RoboDK station: RobodkBasico-2.rdk

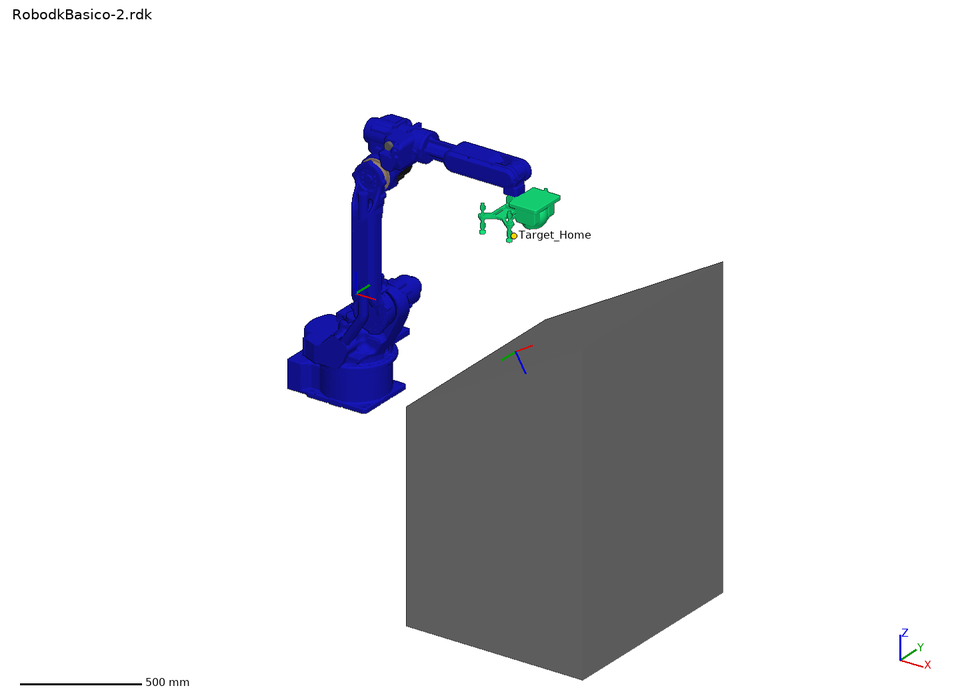
[picture v0: the station drawn from its stored meshes, robots at their saved joint values, targets as dots, program paths as lines]
Station RobodkBasico-2 (saved by RoboDK 6.0.6). Poses are relative to the parent item; angles as X-Y-Z fixed-axis rotations.
Station parameters (name, value as stored): LIN64
  - frame Motoman MH6 Base at (0, 0, 450) mm
    - robot Motoman MH6: 6 axes, payload 6 kg, reach 1422 mm, repeatability 0.08 mm, weight 130 kg
        modified DH rows (alpha deg, a mm, theta deg, d mm): 0, 0, 0, 450; -90, 152, -90, 0; 0, 614, 0, 0; -90, 155, 0, 640; 90, 0, 90, 0; -90, 0, 0, 95
        base shift (0, 0, -450) mm
        joint limits [-170, -90, -175, -180, -45, -360] to [170, 155, 250, 180, 225, 360]; home [0, 0, 0, 0, 0, 0]; saved at [0, 0, 0, 0, 0, 0]
      - tool Ventosas, TCP at (0, 0, 190) mm, size 250 x 290 x 148 mm
    - frame Frame_from_Target1 at (823.2, -34.49, -21.13) mm, rotated rx -180 ry -30 rz 0 deg
      - target Target_Home (Cartesian target) at (225.55, -34.49, -453.06) mm, rotated rx 0 ry -30 rz 0 deg; joints [0, 0, 0, 0, 0, 0] of Motoman MH6
  - object CAJA2 at (1600, 500, 300) mm, rotated rx 180 ry 0 rz 0 deg, size 886.4 x 1000 x 1511.7 mm, geometry from CAJA2.stp
  - Python program RosPolar (listed below)
  - Python program Trébol (listed below)
  - Python program Elipse (listed below)

--- Python program RosPolar ---
from robodk.robolink import *    # API para comunicarte con RoboDK
from robodk.robomath import *    # Funciones matemáticas
import math
from matplotlib.textpath import TextPath
from matplotlib.path import Path
#------------------------------------------------
# 1) Conexión a RoboDK e inicialización
#------------------------------------------------
RDK = Robolink()

# Elegir un robot (si hay varios, aparece un popup)
robot = RDK.ItemUserPick("Selecciona un robot", ITEM_TYPE_ROBOT)
if not robot.Valid():
    raise Exception("No se ha seleccionado un robot válido.")

### Conectar al robot físico
##if not robot.Connect():
##    raise Exception("No se pudo conectar al robot. Verifica que esté en modo remoto y que la configuración sea correcta.")
##
### Confirmar conexión
##if not robot.ConnectedState():
##    raise Exception("El robot no está conectado correctamente. Revisa la conexión.")
##
##print("Robot conectado correctamente.")

#------------------------------------------------
# 2) Cargar el Frame (ya existente) donde quieres dibujar
#    Ajusta el nombre si tu Frame se llama diferente
#------------------------------------------------
frame_name = "Frame_from_Target1"
frame = RDK.Item(frame_name, ITEM_TYPE_FRAME)
if not frame.Valid():
    raise Exception(f'No se encontró el Frame "{frame_name}" en la estación.')

target_name = "Target_Home"
target = RDK.Item(target_name , ITEM_TYPE_TARGET)
if not target.Valid():
    print(f"Error: El target '{target_name}' no existe en la estación.")

# Asignamos este frame al robot
robot.setPoseFrame(frame)
# Usamos la herramienta activa
robot.setPoseTool(robot.PoseTool())

# Ajustes de velocidad y blending
robot.setSpeed(300)   # mm/s - Ajusta según necesites
robot.setRounding(5)  # blending (radio de curvatura)

#------------------------------------------------
# 3) Parámetros de la figura (rosa polar)
#------------------------------------------------
num_points = 100      # Cuántos puntos muestreamos (mayor = más suave)
a = 60
b = 6
z_surface = 0          # Z=0 en el plano del frame
z_safe = 50            # Altura segura para aproximarse y salir

path_jose = TextPath((0, 0), "Jose", size=50)
path_leonardo = TextPath((0, -50), "Leonardo", size=50)

path = Path.make_compound_path(path_jose, path_leonardo)
puntos = path.vertices
instrucciones = path.codes

#------------------------------------------------
# 4) Movimiento al centro en altura segura
#------------------------------------------------
# El centro de la rosa (r=0) corresponde a x=0, y=0
robot.MoveJ(target)
robot.MoveJ(transl(0, 0, z_surface - z_safe))

# Bajamos a la "superficie" (Z=0)
robot.MoveL(transl(0, 0, z_surface))

# #------------------------------------------------
# # 5) Dibujar la rosa polar
# #    r = a - b*cos(theta)
# #    x = r*cos(theta), y = r*sin(theta)
# #------------------------------------------------
# # Recorremos theta de 0 a 2*pi (una vuelta completa)
# full_turn = 2*math.pi

# for i in range(num_points+1):
#     # Fracción entre 0 y 1
#     t = i / num_points
#     # Ángulo actual
#     theta = full_turn * t

#     # Calculamos r
#     r = a - b*math.cos(theta)

#     # Convertimos a coordenadas Cartesianas X, Y
#     x = r * math.cos(theta)
#     y = r * math.sin(theta)

#     # Movemos linealmente (MoveL) en el plano del Frame
#     robot.MoveL(transl(x, y, z_surface))

# # Al terminar, subimos de nuevo para no chocar
# robot.MoveL(transl(x, y, z_surface - z_safe))
# robot.MoveL(target)


# #------------------------------------------------
# # 5) Dibujar la elipse
# #    r = ab/sqrt((b*cos(theta))^2 + (a*sin(theta))^2)
# #    x = r*cos(theta), y = r*sin(theta)
# #------------------------------------------------
# # Recorremos theta de 0 a 2*pi (una vuelta completa)
# full_turn = 2*math.pi

# for i in range(num_points+1):
#     # Fracción entre 0 y 1
#     t = i / num_points
#     # Ángulo actual
#     theta = full_turn * t

#     # Calculamos r
#     r = a*b/sqrt((b*math.cos(theta))**2 + (a*math.sin(theta))**2)

#     # Convertimos a coordenadas Cartesianas X, Y
#     x = r * math.cos(theta)
#     y = r * math.sin(theta)

#     # Movemos linealmente (MoveL) en el plano del Frame
#     robot.MoveL(transl(x, y, z_surface))

# # Al terminar, subimos de nuevo para no chocar
# robot.MoveL(transl(x, y, z_surface - z_safe))
# robot.MoveL(target)

#------------------------------------------------
# 5) Dibujar la trebol b lúbulos
#    r = a*cos(b*theta)
#    x = r*cos(theta), y = r*sin(theta)
#------------------------------------------------
# Recorremos theta de 0 a 2*pi (una vuelta completa)
full_turn = 2*math.pi

for i in range(num_points+1):
    # Fracción entre 0 y 1
    t = i / num_points
    # Ángulo actual
    theta = full_turn * t

    # Calculamos r
    r = a*math.cos(b*theta)-math.cos(theta**2)

    # Convertimos a coordenadas Cartesianas X, Y
    x = r * math.cos(theta)
    y = r * math.sin(theta)

    # Movemos linealmente (MoveL) en el plano del Frame
    robot.MoveL(transl(x, y, z_surface))

# Al terminar, subimos de nuevo para no chocar
robot.MoveL(transl(x, y, z_surface - z_safe))
robot.MoveL(target)


robot.MoveL(transl(150,0,0))
robot.MoveL(transl(0,0,z_surface))

for pt, code in zip(puntos, instrucciones):
    x = pt[1]
    y = pt[0]

    if code == 1:
        # Mover por arriba en el aire y bajar el lápiz
        robot.MoveL(transl(x+150, y, z_surface + z_safe))
        robot.MoveL(transl(x+150, y, z_surface))
    else:
        # Trazo continuo de la letra sobre la superficie
        robot.MoveL(transl(x+150, y, z_surface))

robot.MoveL(transl(x, y, z_surface - z_safe))
robot.MoveJ(target)
print(f"¡Figura (rosa polar) completada en el frame '{frame_name}'!")

--- Python program Trébol ---
from robodk.robolink import *    # API para comunicarte con RoboDK
from robodk.robomath import *    # Funciones matemáticas
import math
from matplotlib.textpath import TextPath
from matplotlib.path import Path
#------------------------------------------------
# 1) Conexión a RoboDK e inicialización
#------------------------------------------------
RDK = Robolink()

# Elegir un robot (si hay varios, aparece un popup)
robot = RDK.ItemUserPick("Selecciona un robot", ITEM_TYPE_ROBOT)
if not robot.Valid():
    raise Exception("No se ha seleccionado un robot válido.")

### Conectar al robot físico
##if not robot.Connect():
##    raise Exception("No se pudo conectar al robot. Verifica que esté en modo remoto y que la configuración sea correcta.")
##
### Confirmar conexión
##if not robot.ConnectedState():
##    raise Exception("El robot no está conectado correctamente. Revisa la conexión.")
##
##print("Robot conectado correctamente.")

#------------------------------------------------
# 2) Cargar el Frame (ya existente) donde quieres dibujar
#    Ajusta el nombre si tu Frame se llama diferente
#------------------------------------------------
frame_name = "Frame_from_Target1"
frame = RDK.Item(frame_name, ITEM_TYPE_FRAME)
if not frame.Valid():
    raise Exception(f'No se encontró el Frame "{frame_name}" en la estación.')

target_name = "Target_Home"
target = RDK.Item(target_name , ITEM_TYPE_TARGET)
if not target.Valid():
    print(f"Error: El target '{target_name}' no existe en la estación.")

# Asignamos este frame al robot
robot.setPoseFrame(frame)
# Usamos la herramienta activa
robot.setPoseTool(robot.PoseTool())

# Ajustes de velocidad y blending
robot.setSpeed(300)   # mm/s - Ajusta según necesites
robot.setRounding(5)  # blending (radio de curvatura)

#------------------------------------------------
# 3) Parámetros de la figura (rosa polar)
#------------------------------------------------
num_points = 100      # Cuántos puntos muestreamos (mayor = más suave)
a = 60
b = 6
z_surface = 0          # Z=0 en el plano del frame
z_safe = 50            # Altura segura para aproximarse y salir

path_jose = TextPath((0, 0), "Jose", size=50)
path_leonardo = TextPath((0, -50), "Leonardo", size=50)

path = Path.make_compound_path(path_jose, path_leonardo)
puntos = path.vertices
instrucciones = path.codes


#------------------------------------------------
# 4) Movimiento al centro en altura segura
#------------------------------------------------
# El centro de la rosa (r=0) corresponde a x=0, y=0
robot.MoveJ(target)
robot.MoveJ(transl(0, 0, z_surface - z_safe))

# Bajamos a la "superficie" (Z=0)
robot.MoveL(transl(0, 0, z_surface))

# #------------------------------------------------
# # 5) Dibujar la rosa polar
# #    r = a - b*cos(theta)
# #    x = r*cos(theta), y = r*sin(theta)
# #------------------------------------------------
# # Recorremos theta de 0 a 2*pi (una vuelta completa)
# full_turn = 2*math.pi

# for i in range(num_points+1):
#     # Fracción entre 0 y 1
#     t = i / num_points
#     # Ángulo actual
#     theta = full_turn * t

#     # Calculamos r
#     r = a - b*math.cos(theta)

#     # Convertimos a coordenadas Cartesianas X, Y
#     x = r * math.cos(theta)
#     y = r * math.sin(theta)

#     # Movemos linealmente (MoveL) en el plano del Frame
#     robot.MoveL(transl(x, y, z_surface))

# # Al terminar, subimos de nuevo para no chocar
# robot.MoveL(transl(x, y, z_surface - z_safe))
# robot.MoveL(target)


# #------------------------------------------------
# # 5) Dibujar la elipse
# #    r = ab/sqrt((b*cos(theta))^2 + (a*sin(theta))^2)
# #    x = r*cos(theta), y = r*sin(theta)
# #------------------------------------------------
# # Recorremos theta de 0 a 2*pi (una vuelta completa)
# full_turn = 2*math.pi

# for i in range(num_points+1):
#     # Fracción entre 0 y 1
#     t = i / num_points
#     # Ángulo actual
#     theta = full_turn * t

#     # Calculamos r
#     r = a*b/sqrt((b*math.cos(theta))**2 + (a*math.sin(theta))**2)

#     # Convertimos a coordenadas Cartesianas X, Y
#     x = r * math.cos(theta)
#     y = r * math.sin(theta)

#     # Movemos linealmente (MoveL) en el plano del Frame
#     robot.MoveL(transl(x, y, z_surface))

# # Al terminar, subimos de nuevo para no chocar
# robot.MoveL(transl(x, y, z_surface - z_safe))
# robot.MoveL(target)

#------------------------------------------------
# 5) Dibujar la trebol b lúbulos
#    r = a*cos(b*theta)
#    x = r*cos(theta), y = r*sin(theta)
#------------------------------------------------
# Recorremos theta de 0 a 2*pi (una vuelta completa)
full_turn = 2*math.pi

for i in range(num_points+1):
    # Fracción entre 0 y 1
    t = i / num_points
    # Ángulo actual
    theta = full_turn * t

    # Calculamos r
    r = a*math.cos(b*theta)

    # Convertimos a coordenadas Cartesianas X, Y
    x = r * math.cos(theta)
    y = r * math.sin(theta)

    # Movemos linealmente (MoveL) en el plano del Frame
    robot.MoveL(transl(x, y, z_surface))

# Al terminar, subimos de nuevo para no chocar
robot.MoveL(transl(x, y, z_surface - z_safe))
robot.MoveL(target)


robot.MoveL(transl(150,0,0))
robot.MoveL(transl(0,0,z_surface))

for pt, code in zip(puntos, instrucciones):
    x = pt[1]
    y = pt[0]

    if code == 1:
        # Mover por arriba en el aire y bajar el lápiz
        robot.MoveL(transl(x+150, y, z_surface + z_safe))
        robot.MoveL(transl(x+150, y, z_surface))
    else:
        # Trazo continuo de la letra sobre la superficie
        robot.MoveL(transl(x+150, y, z_surface))

robot.MoveL(transl(x, y, z_surface - z_safe))
robot.MoveJ(target)
print(f"¡Figura (rosa polar) completada en el frame '{frame_name}'!")

--- Python program Elipse ---
from robodk.robolink import *    # API para comunicarte con RoboDK
from robodk.robomath import *    # Funciones matemáticas
import math
from matplotlib.textpath import TextPath
from matplotlib.path import Path
#------------------------------------------------
# 1) Conexión a RoboDK e inicialización
#------------------------------------------------
RDK = Robolink()

# Elegir un robot (si hay varios, aparece un popup)
robot = RDK.ItemUserPick("Selecciona un robot", ITEM_TYPE_ROBOT)
if not robot.Valid():
    raise Exception("No se ha seleccionado un robot válido.")

### Conectar al robot físico
##if not robot.Connect():
##    raise Exception("No se pudo conectar al robot. Verifica que esté en modo remoto y que la configuración sea correcta.")
##
### Confirmar conexión
##if not robot.ConnectedState():
##    raise Exception("El robot no está conectado correctamente. Revisa la conexión.")
##
##print("Robot conectado correctamente.")

#------------------------------------------------
# 2) Cargar el Frame (ya existente) donde quieres dibujar
#    Ajusta el nombre si tu Frame se llama diferente
#------------------------------------------------
frame_name = "Frame_from_Target1"
frame = RDK.Item(frame_name, ITEM_TYPE_FRAME)
if not frame.Valid():
    raise Exception(f'No se encontró el Frame "{frame_name}" en la estación.')

target_name = "Target_Home"
target = RDK.Item(target_name , ITEM_TYPE_TARGET)
if not target.Valid():
    print(f"Error: El target '{target_name}' no existe en la estación.")

# Asignamos este frame al robot
robot.setPoseFrame(frame)
# Usamos la herramienta activa
robot.setPoseTool(robot.PoseTool())

# Ajustes de velocidad y blending
robot.setSpeed(300)   # mm/s - Ajusta según necesites
robot.setRounding(5)  # blending (radio de curvatura)

#------------------------------------------------
# 3) Parámetros de la figura (rosa polar)
#------------------------------------------------
num_points = 100      # Cuántos puntos muestreamos (mayor = más suave)
a = 40
b = 20
z_surface = 0          # Z=0 en el plano del frame
z_safe = 50            # Altura segura para aproximarse y salir

path_jose = TextPath((0, 0), "Jose", size=50)
path_leonardo = TextPath((0, -50), "Leonardo", size=50)

path = Path.make_compound_path(path_jose, path_leonardo)
puntos = path.vertices
instrucciones = path.codes


#------------------------------------------------
# 4) Movimiento al centro en altura segura
#------------------------------------------------
# El centro de la rosa (r=0) corresponde a x=0, y=0
robot.MoveJ(target)
robot.MoveJ(transl(0, 0, z_surface - z_safe))

# Bajamos a la "superficie" (Z=0)
robot.MoveL(transl(0, 0, z_surface))

# #------------------------------------------------
# # 5) Dibujar la rosa polar
# #    r = a - b*cos(theta)
# #    x = r*cos(theta), y = r*sin(theta)
# #------------------------------------------------
# # Recorremos theta de 0 a 2*pi (una vuelta completa)
# full_turn = 2*math.pi

# for i in range(num_points+1):
#     # Fracción entre 0 y 1
#     t = i / num_points
#     # Ángulo actual
#     theta = full_turn * t

#     # Calculamos r
#     r = a - b*math.cos(theta)

#     # Convertimos a coordenadas Cartesianas X, Y
#     x = r * math.cos(theta)
#     y = r * math.sin(theta)

#     # Movemos linealmente (MoveL) en el plano del Frame
#     robot.MoveL(transl(x, y, z_surface))

# # Al terminar, subimos de nuevo para no chocar
# robot.MoveL(transl(x, y, z_surface - z_safe))
# robot.MoveL(target)


#------------------------------------------------
# 5) Dibujar la elipse
#    r = ab/sqrt((b*cos(theta))^2 + (a*sin(theta))^2)
#    x = r*cos(theta), y = r*sin(theta)
#------------------------------------------------
# Recorremos theta de 0 a 2*pi (una vuelta completa)
full_turn = 2*math.pi

for i in range(num_points+1):
    # Fracción entre 0 y 1
    t = i / num_points
    # Ángulo actual
    theta = full_turn * t

    # Calculamos r
    r = a*b/sqrt((b*math.cos(theta))**2 + (a*math.sin(theta))**2)

    # Convertimos a coordenadas Cartesianas X, Y
    x = r * math.cos(theta)
    y = r * math.sin(theta)

    # Movemos linealmente (MoveL) en el plano del Frame
    robot.MoveL(transl(x, y, z_surface))

# Al terminar, subimos de nuevo para no chocar
robot.MoveL(transl(x, y, z_surface - z_safe))
robot.MoveL(target)

robot.MoveL(transl(150,0,0))
robot.MoveL(transl(0,0,z_surface))

for pt, code in zip(puntos, instrucciones):
    x = pt[1]
    y = pt[0]

    if code == 1:
        # Mover por arriba en el aire y bajar el lápiz
        robot.MoveL(transl(x+150, y, z_surface + z_safe))
        robot.MoveL(transl(x+150, y, z_surface))
    else:
        # Trazo continuo de la letra sobre la superficie
        robot.MoveL(transl(x+150, y, z_surface))

robot.MoveL(transl(x, y, z_surface - z_safe))
robot.MoveJ(target)
print(f"¡Figura (rosa polar) completada en el frame '{frame_name}'!")
